Fanuc KAREL source: KB00009.KL

PROGRAM KB00009
%NOLOCKGROUP
VAR
  P1: REAL
  P2: REAL
  RESULT: REAL
BEGIN
  P1 = 1.0
  P2 = 1.0
  RESULT = ATAN2(P1, P2)
END KB00009
